Fanuc KAREL source: kd00021.compact.KL

PROGRAM KD00021
%STACKSIZE=65535
%PRIORITY=65535
%NOLOCKGROUP
VAR
I : INTEGER
J : INTEGER
B : BOOLEAN
R : REAL
S : STRING[80]
EXTVAL FROM KD00001 : INTEGER
BEGIN
I=EXTVAL
END KD00021
